(* IEC 61131-3 sources: TetherPLC/tests/compat (part 5) *)

(* ---- tc3_mll_case.st ---- *)
// tc3_mll_case.st — Tc3_MLL e2e: simulation-mode linear
// inference, engine-absent error path, and input validation.
PROGRAM tc3_mll_case
VAR
    mask AT %QD0 : UDINT;
    pred : FB_MllPrediction;
    st : INT;
END_VAR
    IF st = 0 THEN
        mask := 0;
        pred.Execute := FALSE;
        // y = 2*x0 + 3*x1 - 1 ; x=(4,5) -> 22
        pred.InputCount := 2;
        pred.X0 := 4.0; pred.X1 := 5.0;
        pred.W0 := 2.0; pred.W1 := 3.0;
        pred.Bias := -1.0;
        pred.FmtIn := 1; pred.FmtOut := 1;   // f32/f32 preferred
        st := 1;
    ELSIF st = 1 THEN
        pred.UseSimulation := TRUE;
        pred.Execute := TRUE;
        st := 2;
    ELSIF st = 2 THEN
        IF pred.YValid AND pred.Y > 21.9 AND pred.Y < 22.1 THEN
            mask := mask OR 1;               // sim inference = 22
            st := 3;
        END_IF;
    ELSIF st = 3 THEN
        pred.Execute := FALSE;
        st := 4;
    ELSIF st = 4 THEN
        IF pred.FmtPreferred THEN
            mask := mask OR 2;               // f32/f32 preferred
            st := 5;
        END_IF;
    ELSIF st = 5 THEN
        pred.UseSimulation := FALSE;
        pred.ModelPath := 'model.onnx';
        pred.Execute := TRUE;                // engine mode, no engine
        st := 6;
    ELSIF st = 6 THEN
        IF pred.Error AND pred.ErrorId = 1 AND NOT pred.YValid THEN
            mask := mask OR 4;               // honest engine-absent
            st := 7;
        END_IF;
    ELSIF st = 7 THEN
        pred.Execute := FALSE;
        st := 8;
    ELSIF st = 8 THEN
        pred.InputCount := 9;                // out of rank range
        pred.Execute := TRUE;
        st := 9;
    ELSIF st = 9 THEN
        IF pred.Error AND pred.ErrorId = 2 THEN
            mask := mask OR 8;
            st := 10;
        END_IF;
    ELSIF st = 10 THEN
        pred.Execute := FALSE;
        st := 11;
    ELSIF st = 11 THEN
        pred.InputCount := 2;
        pred.UseSimulation := FALSE;
        pred.ModelPath := '';                // empty path, engine mode
        pred.Execute := TRUE;
        st := 12;
    ELSIF st = 12 THEN
        IF pred.Error AND pred.ErrorId = 3 THEN
            mask := mask OR 16;
            st := 13;
        END_IF;
    END_IF;

    pred();
END_PROGRAM

(* ---- tc3_nccam_case.st ---- *)
// tc3_nccam_case.st — Tc3_NC_Camming e2e: cam coupling over the
// tplc-motion backend. Master axis runs a velocity move; the slave
// axis is in CSP mode and tracks master*2 through the cam table.
// Also exercises ClearTable and the WritePt point-write edge.
PROGRAM tc3_nccam_case
VAR
    mask   AT %QD0 : DINT;
    st     : INT;
    ax     : FB_MotionAxis;
    axM    : UDINT;
    axS    : UDINT;
    axC    : FB_MotionAxis;   // raw object access for the case
    cpl    : FB_McCamCoupling;
    wrSt   : INT;
    wrN    : INT;
    mPos   : DINT;
    sPos   : DINT;
END_VAR

// ---- st=0: create the two axes ----
IF st = 0 THEN
    mask := 0;
    wrSt := 0;
    wrN := 0;
    ax.UNITS_PER_REV := 1000;
    ax.MAX_VEL := 4000;
    ax.MAX_ACCEL := 20000;
    ax.MAX_DECEL := 20000;
    ax.POS_MIN := -100000;
    ax.POS_MAX := 100000;
    ax.HOME_OFFSET := 0;
    ax.FOLLOW_WINDOW := 10;
    ax.FLAGS := 1;
    ax.OP := 1; ax();
    IF ax.AXIS <> 0 THEN axM := ax.AXIS; END_IF;
    ax.OP := 1; ax();
    IF ax.AXIS <> 0 THEN axS := ax.AXIS; END_IF;
    IF axM <> 0 AND axS <> 0 THEN mask := mask + 1; END_IF;
    st := 1;
END_IF;

// ---- st=1: enable both axes (controlword 0x000F) ----
IF st = 1 THEN
    axC.AXIS := axM;
    axC.OP := 5; axC.INDEX := 16#6040; axC.VALUE := 16#000F; axC();
    axC.AXIS := axS;
    axC.OP := 5; axC.INDEX := 16#6040; axC.VALUE := 16#000F; axC();
    st := 2;
END_IF;

// ---- st=2: slave into CSP mode (0x6060=8) ----
IF st = 2 THEN
    axC.AXIS := axS;
    axC.OP := 5; axC.INDEX := 16#6060; axC.VALUE := 8; axC();
    st := 3;
END_IF;

// ---- st=3: load the cam table directly into the member arrays ----
IF st = 3 THEN
    cpl.MasterPosT[0] := 0.0;    cpl.SlavePosT[0] := 0.0;
    cpl.MasterPosT[1] := 1000.0; cpl.SlavePosT[1] := 2000.0;
    cpl.MasterPosT[2] := 2000.0; cpl.SlavePosT[2] := 4000.0;
    cpl.TableCount := 3;
    IF cpl.TableCountOut = 3 THEN
        mask := mask + 2;      // bit1: table loaded (3 pts)
        st := 4;
    END_IF;
END_IF;

// ---- st=4: master velocity move + coupling live ----
IF st = 4 THEN
    // master: PV mode, target velocity 1000 u/s
    axC.AXIS := axM;
    axC.OP := 5; axC.INDEX := 16#6060; axC.VALUE := 3; axC();
    axC.INDEX := 16#60FF; axC.VALUE := 1000; axC();
    cpl.Execute := TRUE;
    cpl.MasterAxis := axM;
    cpl.SlaveAxis := axS;
    cpl.Periodic := FALSE;
    cpl.Invert := FALSE;
    cpl.MasterScaling := 1.0;
    cpl.SlaveScaling := 1.0;
    cpl.MasterOffset := 0.0;
    cpl.SlaveOffset := 0.0;
    st := 5;
END_IF;

// ---- st=5: wait for the master to cross ~1000, verify slave ~= 2x --
IF st = 5 THEN
    axC.AXIS := axM; axC.OP := 4; axC.INDEX := 16#6064; axC();
    mPos := axC.VALUE;
    IF mPos > 1000 AND mPos < 1400 THEN
        axC.AXIS := axS; axC.OP := 4; axC.INDEX := 16#6064; axC();
        sPos := axC.VALUE;
        // slave target = 2*master at write time; allow scan lag
        IF sPos >= 1900 AND sPos <= 2900 THEN
            mask := mask + 4;  // bit2: cam coupling tracks 2x
            st := 6;
        END_IF;
    ELSIF mPos >= 1400 THEN
        st := 90;            // missed window -> fail
    END_IF;
END_IF;

// ---- st=6: enable periodic wrap; master keeps running past 2000 --
IF st = 6 THEN
    cpl.Periodic := TRUE;
    st := 7;
    wrN := 0;
END_IF;
IF st = 7 THEN
    axC.AXIS := axM; axC.OP := 4; axC.INDEX := 16#6064; axC();
    mPos := axC.VALUE;
    IF mPos > 2050 THEN
        axC.AXIS := axS; axC.OP := 4; axC.INDEX := 16#6064; axC();
        sPos := axC.VALUE;
        // wrapped master ~50-200 -> slave ~100-400
        IF sPos >= 0 AND sPos <= 600 THEN
            mask := mask + 8;  // bit3: periodic wrap
            st := 8;
        END_IF;
    ELSIF wrN > 400 THEN
        st := 90;
    ELSE
        wrN := wrN + 1;
    END_IF;
END_IF;

// ---- st=8: stop coupling, clear table ----
IF st = 8 THEN
    cpl.Execute := FALSE;
    cpl.ClearTable := TRUE;
    st := 9;
END_IF;
IF st = 9 THEN
    IF cpl.TableCountOut = 0 THEN
        mask := mask + 16;     // bit4: table cleared
        st := 10;
    END_IF;
END_IF;

// ---- st=10: WritePt edge writes one point ----
IF st = 10 THEN
    cpl.WritePt := FALSE;
    IF wrSt = 0 THEN
        cpl.PtIndex := 4; cpl.PtMaster := 500.0; cpl.PtSlave := 900.0;
        cpl.WritePt := TRUE; wrSt := 1;
    ELSIF wrSt = 1 THEN
        cpl.WritePt := FALSE;
        IF cpl.TableCountOut = 5 AND cpl.SlavePosT[4] = 900.0 THEN
            mask := mask + 32;  // bit5: WritePt edge
            st := 90;
        END_IF;
    END_IF;
END_IF;

IF st = 90 THEN
    // done
END_IF

// coupling inputs must be driven every scan while active
cpl();
END_PROGRAM

(* ---- tc3_pjlink_case.st ---- *)
PROGRAM Tc3PjlinkCase
VAR
    mask      AT %QD0   : DINT;
    st        : INT;
    g         : FB_PJLink;
    g2        : FB_PJLink;
    p         : FB_PJLink_Power;
    i         : FB_PJLink_Input;
    m         : FB_PJLink_Mute;
    pa        : FB_PJLink_Power;
    pf        : FB_PJLink_Power;
END_VAR

// autonomous PJLink sequence against tests/compat/
// pjlink_test_peer.py (TCP 4352). The peer picks its greeting by
// connection count: conns 1-3 `PJLINK 0` (no auth), conn 4
// `PJLINK 1 a1b2c3d4` accepting md5(nonce+"secret"), conn 5
// `PJLINK 1 deadbeef` rejecting every digest, conns 6+ `PJLINK 0`.
// Each state's bExecute is high only while st equals its index,
// giving every FB one rising edge.
g(sHost := '127.0.0.1', nPort := 4352, nCls := 1, sCmd := 'POWR',
  sParam := '?', sPassword := '', bExecute := st = 0,
  tTimeout := T#2S);
p(sHost := '127.0.0.1', nPort := 4352, sPassword := '',
  nMode := 2, bExecute := st = 1, tTimeout := T#2S);
i(sHost := '127.0.0.1', nPort := 4352, sPassword := '',
  nMode := 0, sInput := '31', bExecute := st = 2,
  tTimeout := T#2S);
pa(sHost := '127.0.0.1', nPort := 4352, sPassword := 'secret',
   nMode := 2, bExecute := st = 3, tTimeout := T#2S);
pf(sHost := '127.0.0.1', nPort := 4352, sPassword := 'wrongpass',
   nMode := 2, bExecute := st = 4, tTimeout := T#2S);
m(sHost := '127.0.0.1', nPort := 4352, sPassword := '',
  nMode := 2, bExecute := st = 5, tTimeout := T#2S);
g2(sHost := '127.0.0.1', nPort := 4352, nCls := 1, sCmd := 'XXXX',
   sParam := '?', sPassword := '', bExecute := st = 6,
   tTimeout := T#2S);

IF st = 0 AND g.bDone THEN
    // POWR ? -> "%1POWR=1": value "1", no auth exchange
    IF g.nStatus = 1 AND g.sValue = '1' AND g.nRespCls = 1 AND
       g.nRespCmd = 1347376978 AND g.nValueLen = 1 AND
       NOT g.bAuthed AND g.nErrId = 0 THEN
        mask := mask + 1;
    END_IF;
    st := 1;
ELSIF st = 1 AND p.bDone THEN
    // Power query -> "1"
    IF p.nStatus = 1 AND p.sValue = '1' AND p.nErrId = 0 THEN
        mask := mask + 2;
    END_IF;
    st := 2;
ELSIF st = 2 AND i.bDone THEN
    // INPT 31 -> "OK"
    IF i.nStatus = 1 AND i.sValue = 'OK' AND i.nErrId = 0 THEN
        mask := mask + 4;
    END_IF;
    st := 3;
ELSIF st = 3 AND pa.bDone THEN
    // authed POWR ? (digest accepted) -> AUTHED, value "1"
    IF pa.nStatus = 1 AND pa.sValue = '1' AND pa.bAuthed AND
       pa.nErrId = 0 THEN
        mask := mask + 8;
    END_IF;
    st := 4;
ELSIF st = 4 AND pf.bDone THEN
    // wrong password -> PJLINK ERRA -> STATUS 5 (authfail)
    IF pf.nStatus = 5 AND pf.nErrId = 0 THEN
        mask := mask + 16;
    END_IF;
    st := 5;
ELSIF st = 5 AND m.bDone THEN
    // AVMT ? -> "31" (muted)
    IF m.nStatus = 1 AND m.sValue = '31' AND m.nErrId = 0 THEN
        mask := mask + 32;
    END_IF;
    st := 6;
ELSIF st = 6 AND g2.bDone THEN
    // unknown command -> "%1XXXX=ERR1": PJLink-level error text,
    // transport status still OK
    IF g2.nStatus = 1 AND g2.sValue = 'ERR1' AND g2.nErrId = 0 THEN
        mask := mask + 64;
    END_IF;
    st := 7;
END_IF;

END_PROGRAM

(* ---- tc3_plctest_case.st ---- *)
// tc3_plctest_case.st — e2e for tc3_plctest (TF1140 surface).
// Every command gets its own scan and a following clear scan, so
// the FB's edge detectors (prev = 0) see a fresh request.
PROGRAM tc3_plctest_case
VAR
    tc : FB_TestCase;
    prep : FB_TestPrepBase;
    suite : FB_TestSuite;
    st : INT;
    mask AT %QD0 : UDINT;
    diag AT %QD4 : UDINT;
END_VAR
    IF st = 0 THEN
        mask := 0;
        tc.nCmd := 5;                        // Reset
        st := 1;
    ELSIF st = 1 THEN
        tc.nCmd := 0;
        st := 2;
    // ---- assertions: set / clear pairs ----
    ELSIF st = 2 THEN
        tc.nAssertCmd := 1; tc.bAssertCond := TRUE;
        st := 3;
    ELSIF st = 3 THEN
        tc.nAssertCmd := 0;
        st := 4;
    ELSIF st = 4 THEN
        tc.nAssertCmd := 2; tc.fActual := 5.0; tc.fExpected := 5.0;
        st := 5;
    ELSIF st = 5 THEN
        tc.nAssertCmd := 0;
        st := 6;
    ELSIF st = 6 THEN
        tc.nAssertCmd := 3;
        tc.fActual := 10.05; tc.fExpected := 10.0; tc.fTolerance := 0.1;
        st := 7;
    ELSIF st = 7 THEN
        tc.nAssertCmd := 0;
        st := 8;
    ELSIF st = 8 THEN
        tc.nAssertCmd := 4;
        tc.fActual := 100.5; tc.fExpected := 100.0; tc.fTolerance := 0.01;
        st := 9;
    ELSIF st = 9 THEN
        tc.nAssertCmd := 0;
        st := 10;
    ELSIF st = 10 THEN
        tc.nAssertCmd := 5; tc.fActual := 7.0; tc.fExpected := 3.0;
        st := 11;
    ELSIF st = 11 THEN
        tc.nAssertCmd := 0;
        IF tc.nAssertions = 5 AND tc.nFailures = 0 AND tc.bSucceeded THEN
            mask := mask OR 1;
        END_IF;
        st := 12;
    ELSIF st = 12 THEN
        tc.nAssertCmd := 2; tc.fActual := 1.0; tc.fExpected := 2.0;
        st := 13;
    ELSIF st = 13 THEN
        tc.nAssertCmd := 0;
        IF tc.nAssertions = 6 AND tc.nFailures = 1
           AND NOT tc.bSucceeded THEN
            mask := mask OR 2;
        END_IF;
        st := 14;
    // ---- step control ----
    ELSIF st = 14 THEN
        tc.nCmd := 1;                        // IncStep
        st := 15;
    ELSIF st = 15 THEN
        tc.nCmd := 0;
        IF tc.nStep = 1 THEN mask := mask OR 4; END_IF;
        st := 16;
    ELSIF st = 16 THEN
        tc.nCmd := 2; tc.nStepArg := 10;     // GoToStep 10
        st := 17;
    ELSIF st = 17 THEN
        tc.nCmd := 0;
        IF tc.nStep = 10 THEN mask := mask OR 8; END_IF;
        st := 18;
    ELSIF st = 18 THEN
        tc.nCmd := 3; tc.bStepCond := FALSE; // IncStepIf false -> stay
        st := 19;
    ELSIF st = 19 THEN
        tc.nCmd := 0;
        IF tc.nStep = 10 THEN mask := mask OR 16; END_IF;
        st := 20;
    ELSIF st = 20 THEN
        tc.nCmd := 3; tc.bStepCond := TRUE;  // IncStepIf true -> 11
        st := 21;
    ELSIF st = 21 THEN
        tc.nCmd := 0;
        IF tc.nStep = 11 THEN mask := mask OR 32; END_IF;
        st := 22;
    // ---- prep block ----
    ELSIF st = 22 THEN
        prep.nAssertCmd := 1; prep.bAssertCond := TRUE;
        st := 23;
    ELSIF st = 23 THEN
        prep.nAssertCmd := 0;
        IF prep.nAssertions = 1 AND prep.bSucceeded THEN
            mask := mask OR 64;
        END_IF;
        st := 24;
    // ---- suite aggregation ----
    ELSIF st = 24 THEN
        suite.bCasePassed := TRUE; suite.nCmd := 1;
        st := 25;
    ELSIF st = 25 THEN
        suite.nCmd := 0;
        st := 26;
    ELSIF st = 26 THEN
        suite.bCasePassed := FALSE; suite.nCmd := 1;
        st := 27;
    ELSIF st = 27 THEN
        suite.nCmd := 0;
        IF suite.nTests = 2 AND suite.nPassed = 1
           AND suite.nFailed = 1 AND NOT suite.bAllPassed THEN
            mask := mask OR 128;
        END_IF;
        st := 28;
    END_IF;
    tc(); prep(); suite();
END_PROGRAM

(* ---- tc3_robotics_case.st ---- *)
// tc3_robotics_case.st — mxAutomation/uniVAL surface e2e:
// connect handshake, move-dispatch validation, engine-absent.
PROGRAM tc3_robotics_case
VAR
    mask AT %QD0 : UDINT;
    grp : FB_RobotGroup;
    cmd : FB_RobotCommand;
    st : INT;
END_VAR
    IF st = 0 THEN
        mask := 0;
        grp.Connect := FALSE;
        cmd.Execute := FALSE;
        grp.Controller := 'krc4-cell';
        grp.RobotCount := 1;
        cmd.GroupConnected := FALSE;
        cmd.MoveType := 1;
        cmd.Velocity := 100.0;
        st := 1;
    ELSIF st = 1 THEN
        // move with no group connection -> not-connected guard
        cmd.Execute := TRUE;
        st := 2;
    ELSIF st = 2 THEN
        IF cmd.Error AND cmd.ErrorId = 5 AND NOT cmd.ReachedTarget THEN
            mask := mask OR 1;
            cmd.Execute := FALSE;
            st := 3;
        END_IF;
    ELSIF st = 3 THEN
        grp.Connect := TRUE;
        st := 4;
    ELSIF st = 4 THEN
        IF grp.Busy THEN mask := mask OR 2; END_IF;
        IF grp.Error AND grp.ErrorId = 1 AND NOT grp.Connected THEN
            mask := mask OR 4;      // license/engine absent
            grp.Connect := FALSE;
            st := 5;
        END_IF;
    ELSIF st = 5 THEN
        grp.Controller := '';      // bad address -> param error
        grp.Connect := TRUE;
        st := 6;
    ELSIF st = 6 THEN
        IF grp.Error AND grp.ErrorId = 2 THEN
            mask := mask OR 8;
            grp.Connect := FALSE;
            st := 7;
        END_IF;
    ELSIF st = 7 THEN
        // connected-flag simulated high -> engine-absent path
        cmd.GroupConnected := TRUE;
        cmd.MoveType := 2;
        cmd.X := 100.0; cmd.Y := 0.0; cmd.Z := 50.0;
        cmd.Execute := TRUE;
        st := 8;
    ELSIF st = 8 THEN
        IF cmd.Error AND cmd.ErrorId = 1 AND NOT cmd.ReachedTarget THEN
            mask := mask OR 16;
            cmd.Execute := FALSE;
            st := 9;
        END_IF;
    ELSIF st = 9 THEN
        cmd.MoveType := 9;         // invalid move -> param error
        cmd.Execute := TRUE;
        st := 10;
    ELSIF st = 10 THEN
        IF cmd.Error AND cmd.ErrorId = 3 THEN
            mask := mask OR 32;
            st := 11;
        END_IF;
    END_IF;

    grp();
    cmd();
END_PROGRAM

(* ---- tc3_rtmon_case.st ---- *)
PROGRAM Tc3RtmonCase
VAR
    mask      AT %QD0   : DINT;
    st        : INT;
    scan_n    : UDINT;
    mkBase    : FB_RTMon_LogMarkBase;
    mkEx      : FB_RTMon_LogMarkBaseEx;
    mStart    : FB_RTMon_LogStart;
    mPlain    : FB_RTMon_LogMark;
    cc        : FB_RtMon;
    c0        : FB_RtMon;
    g0        : FB_RtMon;
    g3        : FB_RtMon;
    g4        : FB_RtMon;
END_VAR

// autonomous realtime-monitor sequence against the tplc-rtmon ring:
// mark x4 (base, ex, simple start, simple plain) -> count=4 ->
// get[0] -> get[3] -> get[4] out-of-range -> clear -> count=0.
mkBase(bExecute := st = 0, nContextId := 1, nGroupId := 10,
       nEventId := 20, nMarkCtrl := 16#E8000000);
mkEx(bExecute := st = 1, nContextId := 2, nGroupId := 30,
     nEventId := 40, nMarkCtrl := 16#60000000);
mStart(bExecute := st = 2, nContextId := 3, bLogCallingTask := TRUE,
       nGroupId := 50, nEventId := 60);
mPlain(bExecute := st = 3, nContextId := 4, bLogCallingTask := FALSE,
       nGroupId := 70, nEventId := 80);

cc.OP := 2;
cc.EXEC := (st = 4) OR (st = 9);
cc();
c0.OP := 4;
c0.EXEC := st = 8;
c0();
g0.OP := 3;
g0.AUX := 0;
g0.EXEC := st = 5;
g0();
g3.OP := 3;
g3.AUX := 3;
g3.EXEC := st = 6;
g3();
g4.OP := 3;
g4.AUX := 4;
g4.EXEC := st = 7;
g4();

IF st = 0 AND mkBase.bDone THEN
    IF mkBase.bError = FALSE AND mkBase.hrErrorCode = 0 THEN
        mask := mask + 1;
    END_IF;
    st := 1;
ELSIF st = 1 AND mkEx.bDone THEN
    IF mkEx.bError = FALSE AND mkEx.hrErrorCode = 0 THEN
        mask := mask + 2;
    END_IF;
    st := 2;
ELSIF st = 2 AND mStart.bDone THEN
    IF mStart.bError = FALSE AND mStart.hrErrorCode = 0 THEN
        mask := mask + 4;
    END_IF;
    st := 3;
ELSIF st = 3 AND mPlain.bDone THEN
    IF mPlain.bError = FALSE AND mPlain.hrErrorCode = 0 THEN
        mask := mask + 8;
    END_IF;
    st := 4;
ELSIF st = 4 AND cc.DONE THEN
    IF cc.RESULT = 4 AND cc.ERRID = 0 THEN
        mask := mask + 16;
    END_IF;
    st := 5;
ELSIF st = 5 AND g0.DONE THEN
    IF g0.ERRID = 0 AND g0.CONTEXT = 1 AND g0.GROUP = 10 AND
       g0.EVENT = 20 AND g0.MARKCTRL = 16#E8000000 THEN
        mask := mask + 32;
    END_IF;
    st := 6;
ELSIF st = 6 AND g3.DONE THEN
    IF g3.ERRID = 0 AND g3.CONTEXT = 4 AND g3.GROUP = 70 AND
       g3.EVENT = 80 AND g3.MARKCTRL = 0 THEN
        mask := mask + 64;
    END_IF;
    st := 7;
ELSIF st = 7 AND g4.DONE THEN
    IF g4.ERRID = 3 THEN
        mask := mask + 128;
    END_IF;
    st := 8;
ELSIF st = 8 AND c0.DONE THEN
    IF c0.ERRID = 0 THEN
        mask := mask + 256;
    END_IF;
    st := 9;
ELSIF st = 9 AND cc.DONE THEN
    IF cc.RESULT = 0 AND cc.ERRID = 0 THEN
        mask := mask + 512;
    END_IF;
    st := 10;
END_IF;

scan_n := scan_n + 1;
END_PROGRAM

(* ---- tc3_s7comm_case.st ---- *)
PROGRAM Tc3S7CommCase
VAR
    mask      AT %QD0   : DINT;
    st        : INT;
    conn      : FB_S7_Connect;
    connBad   : FB_S7_Connect;
    rd        : FB_S7_Read;
    rd2       : FB_S7_Read;
    rd3       : FB_S7_Read;
    wr        : FB_S7_Write;
    rdb       : FB_S7_ReadBit;
    wrb       : FB_S7_WriteBit;
    wdata     : ARRAY[0..239] OF BYTE;
END_VAR

// autonomous S7 sequence against tests/compat/s7_test_peer.py
// (TCP 1102). The peer serves DB1 (256B pattern (i*7+3)) and MK
// area 0 (128B pattern 0xA0+(i&15)) with spec bit semantics.
// Each state's bExecute is high only while st equals its index,
// giving every FB one rising edge; bDone advances the machine.
wdata[0] := 16#DE; wdata[1] := 16#AD;
wdata[2] := 16#BE; wdata[3] := 16#EF;

conn(sHost := '127.0.0.1', nPort := 1102, nRack := 0, nSlot := 2,
     bExecute := st = 0, bClose := st = 8, tTimeout := T#3S);
connBad(sHost := '127.0.0.1', nPort := 19999, nRack := 0, nSlot := 2,
        bExecute := st = 7, bClose := FALSE, tTimeout := T#3S);
rd(nConnHandle := conn.nConnHandle, nArea := 16#84, nDb := 1,
   nByteOff := 10, nLen := 16, bExecute := st = 1,
   tTimeout := T#2S);
wr(nConnHandle := conn.nConnHandle, nArea := 16#84, nDb := 1,
   nByteOff := 0, nLen := 4, pData := wdata, bExecute := st = 2,
   tTimeout := T#2S);
rd2(nConnHandle := conn.nConnHandle, nArea := 16#84, nDb := 1,
    nByteOff := 0, nLen := 4, bExecute := st = 3,
    tTimeout := T#2S);
rdb(nConnHandle := conn.nConnHandle, nArea := 16#83, nDb := 0,
    nByteOff := 5, nBitNo := 0, bExecute := st = 4,
    tTimeout := T#2S);
wrb(nConnHandle := conn.nConnHandle, nArea := 16#83, nDb := 0,
    nByteOff := 5, nBitNo := 1, nBitValue := 1, bExecute := st = 5,
    tTimeout := T#2S);
rd3(nConnHandle := conn.nConnHandle, nArea := 16#84, nDb := 99,
    nByteOff := 0, nLen := 4, bExecute := st = 6,
    tTimeout := T#2S);

IF st = 0 AND conn.bDone THEN
    // connect -> handshake completes, handle issued
    IF conn.nStatus = 1 AND conn.nConnHandle <> 0 AND
       conn.nErrId = 0 THEN
        mask := mask + 1;
    END_IF;
    st := 1;
ELSIF st = 1 AND rd.bDone THEN
    // DB1[10..25] = pattern (i*7+3): first byte 0x49
    IF rd.nStatus = 1 AND rd.nDataLen = 16 AND rd.pData[0] = 16#49
       AND rd.nItemRc = 16#FF AND rd.nErrId = 0 THEN
        mask := mask + 2;
    END_IF;
    st := 2;
ELSIF st = 2 AND wr.bDone THEN
    // write DE AD BE EF -> DB1[0..3]
    IF wr.nStatus = 1 AND wr.nItemRc = 16#FF AND wr.nErrId = 0 THEN
        mask := mask + 4;
    END_IF;
    st := 3;
ELSIF st = 3 AND rd2.bDone THEN
    // readback -> DE AD BE EF
    IF rd2.nStatus = 1 AND rd2.nDataLen = 4 AND
       rd2.pData[0] = 16#DE AND rd2.pData[1] = 16#AD AND
       rd2.pData[2] = 16#BE AND rd2.pData[3] = 16#EF THEN
        mask := mask + 8;
    END_IF;
    st := 4;
ELSIF st = 4 AND rdb.bDone THEN
    // MK5 = 0xA5, bit0 = 1
    IF rdb.nStatus = 1 AND rdb.nBitValue = 1 AND rdb.nErrId = 0 THEN
        mask := mask + 16;
    END_IF;
    st := 5;
ELSIF st = 5 AND wrb.bDone THEN
    // set MK5 bit1 (0xA5 -> 0xA7)
    IF wrb.nStatus = 1 AND wrb.nItemRc = 16#FF AND wrb.nErrId = 0 THEN
        mask := mask + 32;
    END_IF;
    st := 6;
ELSIF st = 6 AND rd3.bDone THEN
    // DB99 unregistered -> item rc 0x0A -> status 5 (s7err)
    IF rd3.nStatus = 5 AND rd3.nItemRc = 16#0A THEN
        mask := mask + 64;
    END_IF;
    st := 7;
ELSIF st = 7 AND connBad.bDone THEN
    // connect to closed port -> conn status 2 (error)
    IF connBad.nStatus = 2 AND connBad.nConnHandle <> 0 THEN
        mask := mask + 128;
    END_IF;
    st := 8;
ELSIF st = 8 THEN
    // bClose := st = 8 gives one rising edge -> session closed
    IF conn.nConnHandle = 0 THEN
        mask := mask + 256;
        st := 9;
    END_IF;
END_IF;

END_PROGRAM

(* ---- tc3_sacn_case.st ---- *)
PROGRAM Tc3SacnCase
VAR
    mask      AT %QD0   : DINT;
    st        : INT;
    inited    : BOOL;
    src       : FB_sACN_Source;
    rcv       : FB_sACN_Receiver;
    hil       : FB_UINT_TO_HighLowArr;
    pair      : ARRAY[1..2] OF BYTE;
    cid       : ARRAY[0..15] OF BYTE;
    dmx       : ARRAY[0..511] OF BYTE;
    dropped0  : ULINT;
END_VAR

IF NOT inited THEN
    inited := TRUE;
    dmx[0] := 16#AA;
    dmx[1] := 16#55;
    dmx[2] := 16#01;
    dmx[3] := 16#02;
END_IF;

// source: universe 1, priority 100, 50 ms interval, auto CID
src(bEnable := TRUE, nUniverse := 1, nPriority := 100,
    nSyncUniverse := 0, sSourceName := 'SRC1',
    nSendIntervalMs := 50, nTimeToLive := 0,
    bOptionForceSync := FALSE, bOptionStreamTerminated := FALSE,
    bOptionPreviewData := FALSE, nDmxStartCode := 0,
    bSendSync := FALSE, bSendDiscovery := FALSE,
    cid := cid, DmxData := dmx, nDmxLength := 4);

// receiver: universe 1 on the default sACN port
rcv(bEnable := TRUE, nUniverse := 1, nSyncUniverse := 0,
    nPort := 5568);

// phase A: only our source is on the wire -> payload/name/prio
IF st = 0 AND rcv.nDataPackets >= 3 AND rcv.bHaveData THEN
    IF rcv.nDmxLength = 4 AND rcv.DmxData[0] = 16#AA AND
       rcv.DmxData[1] = 16#55 AND rcv.DmxData[2] = 16#01 AND
       rcv.DmxData[3] = 16#02 AND rcv.sSourceName = 'SRC1' AND
       rcv.nPriority = 100 AND rcv.nErrId = 0 THEN
        mask := mask + 1;
    END_IF;
    dropped0 := rcv.nDroppedPackets;
    st := 1;
// phase B: peer's priority-10 HIPRI packet preempts the source
ELSIF st = 1 AND rcv.sSourceName = 'HIPRI' THEN
    IF rcv.nPriority = 10 AND rcv.nDmxLength = 3 AND
       rcv.DmxData[0] = 16#33 AND rcv.DmxData[1] = 16#44 AND
       rcv.DmxData[2] = 16#55 THEN
        mask := mask + 2;
    END_IF;
    st := 2;
// phase C: peer's priority-200 LOWPR and our priority-100 source
// are both dropped once HIPRI holds the channel
ELSIF st = 2 AND rcv.sSourceName = 'HIPRI' AND
          rcv.nDroppedPackets > dropped0 + 1 THEN
    mask := mask + 4;
    st := 3;
// phase D: pure-IEC helpers
ELSIF st = 3 THEN
    pair[1] := 0;
    pair[2] := 1;
    hil(bExecute := TRUE, Value := 16#1234);
    IF F_HighLowArr_TO_UINT(pair) = 1 AND
       F_UNIVERSE_TO_MulticastAdr(1) = 16#EFFF0001 AND
       F_UNIVERSE_TO_MulticastAdr(63999) = 16#EFFFF9FF AND
       hil.bDone AND hil.HighByte = 16#12 AND hil.LowByte = 16#34 THEN
        mask := mask + 8;
        st := 4;
    END_IF;
END_IF;

END_PROGRAM

(* ---- tc3_speech_case.st ---- *)
// tc3_speech_case.st — Tc3_Speech e2e: honest engine-absent
// handshake — TTS/SR commands run Busy for a bounded window then
// fail with ErrorId=1 (engine-unavailable); parameter validation
// fires immediately (ErrorId=2/3).
PROGRAM tc3_speech_case
VAR
    mask AT %QD0 : UDINT;
    tts : FB_TextToSpeech;
    sr : FB_SpeechRecognition;
    st : INT;
END_VAR
    IF st = 0 THEN
        mask := 0;
        tts.Speak := FALSE;
        sr.Listen := FALSE;
        tts.Utterance := 'hello axis';
        tts.ConfigurationId := 1;
        tts.LanguageId := 0;
        sr.ConfigurationId := 1;
        st := 1;
    ELSIF st = 1 THEN
        tts.Speak := TRUE;         // valid command -> handshake
        st := 2;
    ELSIF st = 2 THEN
        IF tts.Busy THEN mask := mask OR 1; END_IF;
        IF tts.Error AND tts.ErrorId = 1 THEN
            mask := mask OR 2;      // engine-unavailable reported
            st := 3;
        END_IF;
    ELSIF st = 3 THEN
        tts.Speak := FALSE;
        st := 4;
    ELSIF st = 4 THEN
        tts.Utterance := '';       // empty -> param error
        tts.Speak := TRUE;
        st := 5;
    ELSIF st = 5 THEN
        IF tts.Error AND tts.ErrorId = 2 THEN
            mask := mask OR 4;      // bad-utterance validated
            st := 6;
        END_IF;
    ELSIF st = 6 THEN
        tts.Speak := FALSE;
        sr.Listen := TRUE;         // valid recognition command
        st := 7;
    ELSIF st = 7 THEN
        IF sr.Error AND sr.ErrorId = 1 AND NOT sr.ResultValid THEN
            mask := mask OR 8;      // SR engine-absent, no fake text
            st := 8;
        END_IF;
    ELSIF st = 8 THEN
        sr.Listen := FALSE;        // let the FB re-arm one scan
        st := 9;
    ELSIF st = 9 THEN
        sr.ConfigurationId := 0;   // missing config -> param error
        sr.Listen := TRUE;
        st := 10;
    ELSIF st = 10 THEN
        IF sr.Error AND sr.ErrorId = 3 THEN
            mask := mask OR 16;
            st := 11;
        END_IF;
    END_IF;

    tts();
    sr();
END_PROGRAM

(* ---- tc3_vision_case.st ---- *)
// tc3_vision_case.st — Tc3_Vision e2e: camera-open handshake,
// acquire-image not-open guard, job dispatch — all honest
// engine-absent paths.
PROGRAM tc3_vision_case
VAR
    mask AT %QD0 : UDINT;
    cam : FB_VN_GevCamera;
    acq : FB_VN_AcquireImage;
    job : FB_VN_JobControl;
    st : INT;
END_VAR
    IF st = 0 THEN
        mask := 0;
        cam.Open := FALSE;
        acq.Trigger := FALSE;
        job.Execute := FALSE;
        acq.CameraOpen := FALSE;
        cam.IpAddress := '192.168.1.10';
        cam.Port := 3956;
        st := 1;
    ELSIF st = 1 THEN
        // acquire with no open channel -> not-open guard
        acq.Trigger := TRUE;
        st := 2;
    ELSIF st = 2 THEN
        IF acq.Error AND acq.ErrorId = 5 AND NOT acq.ImageReady THEN
            mask := mask OR 1;
            acq.Trigger := FALSE;
            st := 3;
        END_IF;
    ELSIF st = 3 THEN
        cam.Open := TRUE;          // valid address -> handshake
        st := 4;
    ELSIF st = 4 THEN
        IF cam.Busy THEN mask := mask OR 2; END_IF;
        IF cam.Error AND cam.ErrorId = 1 AND NOT cam.Opened THEN
            mask := mask OR 4;      // engine-absent on open
            cam.Open := FALSE;
            st := 5;
        END_IF;
    ELSIF st = 5 THEN
        cam.IpAddress := '';       // bad address -> param error
        cam.Open := TRUE;
        st := 6;
    ELSIF st = 6 THEN
        IF cam.Error AND cam.ErrorId = 2 THEN
            mask := mask OR 8;
            cam.Open := FALSE;
            st := 7;
        END_IF;
    ELSIF st = 7 THEN
        job.JobType := 42;         // valid job -> handshake
        job.Execute := TRUE;
        st := 8;
    ELSIF st = 8 THEN
        IF job.Error AND job.ErrorId = 1 AND NOT job.ResultValid THEN
            mask := mask OR 16;
            job.Execute := FALSE;
            st := 9;
        END_IF;
    ELSIF st = 9 THEN
        job.JobType := 0;          // bad job id -> param error
        job.Execute := TRUE;
        st := 10;
    ELSIF st = 10 THEN
        IF job.Error AND job.ErrorId = 3 THEN
            mask := mask OR 32;
            st := 11;
        END_IF;
    END_IF;

    cam();
    acq();
    job();
END_PROGRAM

(* ---- tc3_xmlsrv_case.st ---- *)
// tc3_xmlsrv_case.st — e2e for tc3_xmlsrv (file-backed XML store).
PROGRAM tc3_xmlsrv_case
VAR
    wr : FB_XmlSrvWrite;
    rd : FB_XmlSrvRead;
    wrn : FB_XmlSrvWriteByName;
    rdn : FB_XmlSrvReadByName;
    obf : FB_XmlSrvIsObfuscationEnabled;
    st : INT;
    mask AT %QD0 : UDINT;
    diag AT %QD4 : UDINT;
END_VAR
    diag := st;
    IF st = 0 THEN
        mask := 0;
        wr.sFilePath := '/tmp/tplc_xmlsrv_e2e.xml';
        wr.sXPath := 'PLC/Tags/Temperature';
        wr.sValue := '21.5';
        wr.bExecute := TRUE;
        st := 1;
    ELSIF st = 1 THEN
        IF wr.bDone THEN mask := mask OR 1; END_IF;
        wr.bExecute := FALSE;
        rd.sFilePath := '/tmp/tplc_xmlsrv_e2e.xml';
        rd.sXPath := 'PLC/Tags/Temperature';
        st := 2;
    ELSIF st = 2 THEN
        rd.bExecute := TRUE;
        st := 3;
    ELSIF st = 3 THEN
        IF NOT rd.bError AND FIND(rd.sValue, '21.5') = 1 THEN
            mask := mask OR 2;
        END_IF;
        rd.bExecute := FALSE;
        // second element via the ByName variant
        wrn.sFilePath := '/tmp/tplc_xmlsrv_e2e.xml';
        wrn.sXPath := 'PLC/Tags/Pressure';
        wrn.sValue := '7.25';
        st := 4;
    ELSIF st = 4 THEN
        wrn.bExecute := TRUE;
        st := 5;
    ELSIF st = 5 THEN
        IF wrn.bDone THEN mask := mask OR 4; END_IF;
        wrn.bExecute := FALSE;
        rdn.sFilePath := '/tmp/tplc_xmlsrv_e2e.xml';
        rdn.sXPath := 'PLC/Tags/Pressure';
        st := 6;
    ELSIF st = 6 THEN
        rdn.bExecute := TRUE;
        st := 7;
    ELSIF st = 7 THEN
        IF NOT rdn.bError AND FIND(rdn.sValue, '7.25') = 1 THEN
            mask := mask OR 8;
        END_IF;
        rdn.bExecute := FALSE;
        // first element must still be intact after the rewrite
        rd.sXPath := 'PLC/Tags/Temperature';
        st := 8;
    ELSIF st = 8 THEN
        rd.bExecute := TRUE;
        st := 9;
    ELSIF st = 9 THEN
        IF NOT rd.bError AND FIND(rd.sValue, '21.5') = 1 THEN
            mask := mask OR 16;
        END_IF;
        rd.bExecute := FALSE;
        // missing key -> error
        rd.sXPath := 'PLC/Tags/Absent';
        st := 10;
    ELSIF st = 10 THEN
        rd.bExecute := TRUE;
        st := 11;
    ELSIF st = 11 THEN
        IF rd.bError THEN mask := mask OR 32; END_IF;
        rd.bExecute := FALSE;
        obf.bExecute := TRUE;
        st := 12;
    ELSIF st = 12 THEN
        IF obf.bDone AND NOT obf.bEnabled THEN mask := mask OR 64; END_IF;
        obf.bExecute := FALSE;
        st := 13;
    END_IF;
    wr(); rd(); wrn(); rdn(); obf();
END_PROGRAM
